// TIA Portal V21 export
// export: Created 2000-01-01T00:00:00.0000000Z, ExportSetting None
TYPE "UDT_HMI_ButtonDebounce"
   STRUCT
      bHmiToggleCmd { ExternalWritable := 'False'} : Bool;   // HMI软按钮翻转触发
      bHmiForceOn { ExternalWritable := 'False'} : Bool;   // HMI强制置位开机
      bHmiForceOff { ExternalWritable := 'False'} : Bool;   // HMI强制复位关机
      tDebounceTime { ExternalWritable := 'False'} : Time;   // 防抖延时时间设定（默认 T#50ms）
      tElapsedMs { ExternalWritable := 'False'} : DInt;   // 内部保持：当前防抖累计毫秒数
      bDebouncedState { ExternalWritable := 'False'} : Bool;   // 状态反馈：防抖后的稳定按钮状态
      bPrevDebounced { ExternalWritable := 'False'} : Bool;   // 内部保持：上一周期防抖状态（用于取沿）
      bToggleOut { ExternalWritable := 'False'} : Bool;   // 状态反馈：当前单键启停翻转锁存输出
      wStatus { ExternalWritable := 'False'} : Word;   // 状态码：16#0000正常, 16#8401急停强制释放
   END_STRUCT;
END_TYPE
